(* IEC 61131-3 sources: iecf/crates/iecf-syntax/tests/corpus, 7 files *)

(* ---- demo_globals.gvl ---- *)
(* demo_globals.gvl - the project's plain globals (CODESYS's GVL).
   The build puts these blocks into the CONFIGURATION and gives every
   POU that uses one its VAR_EXTERNAL (spec/io-tags.md §7). *)
VAR_GLOBAL
    counter : INT;
    top_value : INT := 100;   (* counter wraps past this *)
    speed : REAL := 1.5;
END_VAR
VAR_GLOBAL CONSTANT
    increment : INT := 3;
END_VAR
VAR_GLOBAL RETAIN
    total : DINT;             (* survives an online change *)
END_VAR

(* ---- core.st ---- *)
(* One of each Ed.2 core construct the Prokop examples do not use. *)
TYPE
    RunMode : (Idle, Running, Fault) := Idle;
    Level : INT (0..100) := 50;
    Code : UINT (Ok := 0, Warn := 1, Bad := 2);
    Point : STRUCT
        x : REAL;
        y : REAL := 1.5;
    END_STRUCT;
    Row : ARRAY [1..3] OF INT := [1, 2, 3];
    Name : STRING[20] := 'none';
END_TYPE

FUNCTION Clamp : INT
VAR_INPUT
    v, lo, hi : INT;
END_VAR
IF v < lo THEN
    Clamp := lo;
ELSIF v > hi THEN
    Clamp := hi;
ELSE
    Clamp := v;
END_IF;
END_FUNCTION

FUNCTION_BLOCK Ctr
VAR_INPUT
    pulse : BOOL R_EDGE;
    reset : BOOL;
END_VAR
VAR_OUTPUT
    count : DINT;
END_VAR
VAR_IN_OUT
    total : LINT;
END_VAR
VAR_TEMP
    inc : DINT := 1;
END_VAR
IF reset THEN
    count := 0;
    RETURN;
END_IF;
IF pulse THEN
    count := count + inc;
    total := total + 1;
END_IF;
END_FUNCTION_BLOCK

PROGRAM core
VAR
    mode : RunMode;
    grid : ARRAY [0..2, 0..2] OF REAL := [9(0.0)];
    p : Point := (x := 1.0, y := 2.0);
    c : Ctr;
    big : LINT;
    i, n : INT;
    w : WORD := 16#00FF;
    b : BYTE := 2#1010_0101;
    s : STRING := 'it$'s $$5$N';
    ws : WSTRING := "wide$0041";
    t : TIME := T#1h2m3s4ms;
    d : DATE := D#2026-11-05;
    tod_v : TOD := TOD#12:00:00.5;
    dt_v : DT := DT#2026-11-05-12:00:00;
    r : REAL := -1.5E-3;
    ok : BOOL;
    flag : BOOL := BOOL#TRUE;
    neg : INT := INT#-5;
END_VAR
VAR CONSTANT
    MAX_N : INT := 10;
END_VAR

CASE mode OF
    Idle:
        mode := Running;
    Running, Fault:
        ;
END_CASE;

CASE i OF
    1, 2..5: n := 1;
    -1: n := -1;
ELSE
    n := 0;
END_CASE;

FOR i := 0 TO 2 BY 1 DO
    grid[i, i] := 1.0;
    IF i = MAX_N THEN
        EXIT;
    END_IF;
END_FOR;

WHILE n < MAX_N DO
    n := n + 1;
    IF n MOD 2 = 0 THEN
        CONTINUE;
    END_IF;
END_WHILE;

REPEAT
    n := n - 1;
UNTIL n <= 0
END_REPEAT;

c(pulse := ok, reset := FALSE, count => big, total := big);
n := Clamp(v := n, lo := 0, hi := MAX_N);
n := Clamp(n, 0, MAX_N);
ok := NOT ok AND (n > 0 OR n < -2) XOR w.3;
r := -2.0 ** 2.0 + p.x * 3.0 / 2.0;
mode := RunMode#Fault;
END_PROGRAM

(* ---- demo_fb_aux.st ---- *)
(* demo_fb_aux.st - exercises the aux region (spec/abi.md §5a,
 * Prokop's toolchain): a real TON timer's public interface members
 * (IN/PT/Q/ET) and a plain top-level PROGRAM-local variable, both
 * non-located and non-retained, so neither the process image nor the
 * retain region would expose them without the aux bridge.
 *
 * VAR blocks are deliberately split (FB instance declarations separate
 * from the AT-located one): mixing them in one VAR block is refused
 * (PROPOSAL.md §1e).
 *)
PROGRAM main
VAR
    fill_tmr : TON;
END_VAR
VAR
    start_pb AT %IX0.0 : BOOL;
END_VAR
VAR
    local_counter : INT;
END_VAR
fill_tmr(IN := start_pb, PT := T#20s);
local_counter := local_counter + 1;
END_PROGRAM

CONFIGURATION Config0
    RESOURCE Res0 ON PLC
        TASK task0(INTERVAL := T#10ms, PRIORITY := 0);
        PROGRAM instance0 WITH task0 : main;
    END_RESOURCE
END_CONFIGURATION

(* ---- demo_ld.st ---- *)
(* demo_ld.st - a LADDER diagram through the full pipeline, exactly as the
 * graphical path produces it (spec/graphical-languages.md §2, §8 G4): the
 * POU below is byte-for-byte what the Workbench emits for the ladder in
 * workbench/src/lib/graphical/fbd-ladder.test.ts ("demo ladder parity"
 * guards the match), and the CONFIGURATION mirrors what the server
 * generates from prokop.json.
 *
 * LD is not a textual language - it is FBD plus three element
 * types (PLCopen says so literally: LD = commonObjects + fbdObjects +
 * ldObjects), compiled by the SAME graph->ST generator. What the rungs say:
 *
 *   |--| |--+--|/|--( )--    seal-in latch: start OR motor, AND NOT halt
 *   |  start|  halt  motor
 *   |--| |--+
 *   |  motor
 *
 *   |--|P|----------( )--    a rising-edge contact: one scan per press,
 *   |   jog         pulsed   via the R_TRIG the generator synthesized
 *
 * Note the rail contributes nothing to the expression (`AND(TRUE, x)` is
 * just `x`) and the edge trigger is called BEFORE the rungs: IEC's |P|
 * fires on an edge of the CONTACT's variable, never of the rung.
 *)
PROGRAM Latch
VAR
    start AT %IX0.0 : BOOL;
    halt AT %IX0.1 : BOOL;
    jog AT %IX0.2 : BOOL;
    motor AT %QX0.0 : BOOL;
    pulsed AT %QX0.1 : BOOL;
END_VAR
VAR
    RTRIG_C4 : R_TRIG;
END_VAR

RTRIG_C4(CLK := jog);
motor := AND(OR(start, motor), NOT(halt));
pulsed := RTRIG_C4.Q;

END_PROGRAM

CONFIGURATION Config0
    RESOURCE Res0 ON PLC
        TASK task0(INTERVAL := T#10ms, PRIORITY := 0);
        PROGRAM instance0 WITH task0 : Latch;
    END_RESOURCE
END_CONFIGURATION

(* ---- demo_sfc.st ---- *)
(* demo_sfc.st - textual SFC through the full pipeline, exactly as the
 * graphical path produces it (spec/graphical-languages.md §3): the POU
 * below is byte-for-byte what the Workbench's SFC generator emits for
 * the demo chart in workbench/src/lib/graphical/sfc-generate.test.ts
 * ("demo chart parity" test guards the match - edit either side and
 * that test fails), and the CONFIGURATION mirrors what the server
 * generates from prokop.json. The SFC is compiled as SFC, not turned
 * into ST first.
 *)
PROGRAM DemoSfc
VAR
    start AT %IX0.0 : BOOL;
    running AT %QX0.0 : BOOL;
    entries AT %QW1 : INT;
END_VAR

INITIAL_STEP Idle:
    IdleMode(N);
END_STEP

STEP Active:
    ActiveMode(N);
    EntryCount(P);
END_STEP

TRANSITION FROM Idle TO Active
    := start;
END_TRANSITION

TRANSITION FROM Active TO Idle
    := NOT start;
END_TRANSITION

ACTION IdleMode:
    running := FALSE;
END_ACTION

ACTION ActiveMode:
    running := TRUE;
END_ACTION

ACTION EntryCount:
    entries := entries + 1;
END_ACTION

END_PROGRAM

CONFIGURATION Config0
    RESOURCE Res0 ON PLC
        TASK task0(INTERVAL := T#10ms, PRIORITY := 0);
        PROGRAM instance0 WITH task0 : DemoSfc;
    END_RESOURCE
END_CONFIGURATION

(* ---- demo_switch.st ---- *)
(* demo_switch.st - Prokop's first spike (ARCHITECTURE.md §13): a real ST
 * program, compiled by a real IEC compiler, run through the real toolchain
 * pipeline into a module a real scan engine loads and executes.
 *
 * A seal-in latch plus a pass-through on located I/O (exercises
 * the toolchain's process-image binding), plus a VAR RETAIN counter and
 * totalizer (exercises the toolchain's bridge to spec/abi.md §5's retain
 * region, see toolchain/README.md).
 *)
PROGRAM main
VAR
    di0 AT %IX0.0 : BOOL;   (* set: latches dout0 on *)
    di1 AT %IX0.1 : BOOL;   (* set: latches dout0 off *)
    sp AT %IW0 : INT;       (* setpoint in *)
    dout0 AT %QX0.0 : BOOL;
    pv AT %QW0 : INT;       (* setpoint echoed out *)
END_VAR
VAR RETAIN
    scan_counter : DINT;    (* must survive an online slot swap *)
    totalizer : LREAL;      (* accumulates pv every scan di0 is set *)
END_VAR

IF di0 THEN
    dout0 := TRUE;
    totalizer := totalizer + INT_TO_LREAL(pv);
END_IF;
IF di1 THEN
    dout0 := FALSE;
END_IF;
pv := sp;
scan_counter := scan_counter + 1;

END_PROGRAM

CONFIGURATION Config0
    RESOURCE Res0 ON PLC
        TASK task0(INTERVAL := T#10ms, PRIORITY := 0);
        PROGRAM instance0 WITH task0 : main;
    END_RESOURCE
END_CONFIGURATION

(* ---- demo_time_types.st ---- *)
(* demo_time_types.st - TIME, DATE, TOD and DT (spec/abi.md §6),
   arithmetic on them, and RETAIN of a TIME, a STRING and a DATE.

   No variable is called `dt` or `tod`: some compilers reserve the type
   names. *)
PROGRAM main
VAR
    elapsed : TIME := T#1500ms;
    shift_start : TOD := TOD#14:30:15.25;
    stamp : DT := DT#2026-10-04-14:30:15;
    today : DATE := D#2026-10-04;
    half : TIME;
    gap : TIME;
END_VAR
VAR RETAIN
    hold : TIME := T#5s;
    note : STRING := 'kept';
    since : DATE := D#2000-01-01;
    ticks : DINT;
END_VAR
elapsed := elapsed + T#10ms;
shift_start := shift_start + T#1s;
stamp := stamp + T#1s;
half := elapsed / 2;
gap := elapsed - T#500ms;
ticks := ticks + 1;
END_PROGRAM

CONFIGURATION Config0
    RESOURCE Res0 ON PLC
        TASK task0(INTERVAL := T#10ms, PRIORITY := 0);
        PROGRAM instance0 WITH task0 : main;
    END_RESOURCE
END_CONFIGURATION
